(* IEC 61131-3 sources: codesys-framework/txt/application/WeVe Core (library)/10 Mode/FB_Mode/States, 12 files *)

(* ---- HandleEmergencyStop.method.st ---- *)
METHOD PROTECTED HandleEmergencyStop
VAR_INPUT
END_VAR

// --- BEGIN IMPLEMENTATION ---

IF _fbEmergencyStopMod.State = E_EmergencyStopState.NOK THEN

	CASE _eState OF

		E_ModeStates.Invalid : ;
		E_ModeStates.Off,
		E_ModeStates.Initialize,
		E_ModeStates.Standby : _eState := E_ModeStates.Invalid;

		E_ModeStates.Starting,
		E_ModeStates.Run  : _eState := E_ModeStates.QuickStop;

		E_ModeStates.Stop,
		E_ModeStates.Safe,
		E_ModeStates.QuickStop,
		E_ModeStates.Reset : ;

	END_CASE

END_IF

(* ---- ProcessInitialize.method.st ---- *)
METHOD PROTECTED ProcessInitialize
VAR_INPUT
END_VAR
VAR
END_VAR

// --- BEGIN IMPLEMENTATION ---

_iStateStarting := 0;
_iStateRun := 0;
_iStateStop := 0;
_iStateEStop := 0;
_iStateReset := 0;

_eState := E_ModeStates.Standby;

(* ---- ProcessInvalid.method.st ---- *)
METHOD PROTECTED ProcessInvalid
VAR_INPUT
END_VAR

// --- BEGIN IMPLEMENTATION ---

(* ---- ProcessOff.method.st ---- *)
METHOD PROTECTED ProcessOff
VAR_INPUT
END_VAR

// --- BEGIN IMPLEMENTATION ---

IF _xActive THEN
	_eState := E_ModeStates.Initialize;
END_IF

(* ---- ProcessQuickStop.method.st ---- *)
METHOD PROTECTED ProcessQuickStop
VAR_INPUT
END_VAR
VAR
END_VAR

// --- BEGIN IMPLEMENTATION ---

(* ---- ProcessReset.method.st ---- *)
METHOD PROTECTED ProcessReset
VAR_INPUT
END_VAR
VAR
END_VAR

// --- BEGIN IMPLEMENTATION ---

(* ---- ProcessRun.method.st ---- *)
METHOD PROTECTED ProcessRun
VAR_INPUT
END_VAR

// --- BEGIN IMPLEMENTATION ---

(* ---- ProcessSafe.method.st ---- *)
METHOD PROTECTED ProcessSafe
VAR_INPUT
END_VAR

// --- BEGIN IMPLEMENTATION ---

(* ---- ProcessStandby.method.st ---- *)
METHOD PROTECTED ProcessStandby
VAR_INPUT
END_VAR

// --- BEGIN IMPLEMENTATION ---

(* ---- ProcessStarting.method.st ---- *)
METHOD PROTECTED ProcessStarting
VAR_INPUT
END_VAR

// --- BEGIN IMPLEMENTATION ---

(* ---- ProcessStates.method.st ---- *)
METHOD PROTECTED ProcessStates
VAR_INPUT
END_VAR

// --- BEGIN IMPLEMENTATION ---

CASE _eState OF

	E_ModeStates.Off : ProcessOff();
	E_ModeStates.Initialize : ProcessInitialize();
	E_ModeStates.Standby : ProcessStandby();
	E_ModeStates.Starting : ProcessStarting();
	E_ModeStates.Run : ProcessRun();
	E_ModeStates.Stop : ProcessStop();
	E_ModeStates.QuickStop : ProcessQuickStop();
	E_ModeStates.Invalid : ProcessInvalid();
	E_ModeStates.Reset : ProcessReset();
	E_ModeStates.Safe : ProcessSafe();

END_CASE

(* ---- ProcessStop.method.st ---- *)
METHOD PROTECTED ProcessStop
VAR_INPUT
END_VAR
VAR
END_VAR

// --- BEGIN IMPLEMENTATION ---
